DATA_BLOCK "FRK_Carriers"
{ S7_Optimized_Access := 'TRUE' }
VERSION : 0.1
NON_RETAIN
VAR
    Slots {ExternalAccessible := 'False'; ExternalVisible := 'False'; ExternalWritable := 'False'} : Array[0..4] of "FRK_Carrier";
END_VAR
BEGIN
END_DATA_BLOCK
